            Waypoint PosA_pick: TCP in base x=15.039 y=-636.805 z=98.001 mm, rx=-1.0907 ry=1.4048 rz=-1.4136 rad; joints [-59.046, -153.942, -49.224, -157.253, 46.333, 1.224] deg
            URCap Gripper (Robotiq_Grippers, Robotiq Inc.) dataModel(position=100.0, force=30.19607843137255, speed=49.80392156862745, positionInDouble=100.0, forceInDouble=30.19607843137255, speedInDouble=49.80392156862745, slaveIds=[9], blocking=true, robotCompliant=false)
            Waypoint PosA_up: motionParameters(jointSpeed=1.047198 jointAcceleration=1.396263 cartesianSpeed=0.04 cartesianAcceleration=0.3); TCP in base x=16.801 y=-634.608 z=234.973 mm, rx=-1.0907 ry=1.4048 rz=-1.4136 rad; joints [-58.842, -146.487, -43.11, -170.828, 46.488, 1.231] deg
            Waypoint Postions_otw: motionParameters(blendRadius=0.01); TCP in base x=-10.897 y=-533.369 z=288.851 mm, rx=-1.2337 ry=1.1953 rz=-1.2073 rad; joints [-51.497, -119.089, -83.078, -158.276, 37.645, 1.224] deg
        ElseIf powder_position≟"Position2"
          MoveJ speed 60 deg/s, acceleration 80 deg/s^2 (useActiveTCP=true optimoveEnabled=false optiMoveSpeed=0.3 optiMoveAcceleration=0.09) feature=Base
            Waypoint Postions_otw: motionParameters(blendRadius=0.01); TCP in base x=-10.897 y=-533.369 z=288.851 mm, rx=-1.2337 ry=1.1953 rz=-1.2073 rad; joints [-51.497, -119.089, -83.078, -158.276, 37.645, 1.224] deg
          URCap Gripper (Robotiq_Grippers, Robotiq Inc.) dataModel(position=0.0, force=30.19607843137255, speed=49.80392156862745, positionInDouble=0.0, forceInDouble=30.19607843137255, speedInDouble=49.80392156862745, slaveIds=[9], blocking=true, robotCompliant=false)
          MoveL speed 250 mm/s, acceleration 1200 mm/s^2 (useActiveTCP=true optimoveEnabled=false optiMoveSpeed=0.3 optiMoveAcceleration=0.09) feature=Base
            Waypoint PosB_up: motionParameters(blendRadius=0.01); TCP in base x=239.473 y=-492.481 z=220.768 mm, rx=-1.2337 ry=1.1953 rz=-1.2073 rad; joints [-33.233, -137.947, -61.305, -161.095, 55.866, 1.01] deg
            Waypoint PosB_pick: TCP in base x=240.63 y=-494.559 z=96.393 mm, rx=-1.2337 ry=1.1953 rz=-1.2073 rad; joints [-33.324, -146.292, -65.182, -148.873, 55.811, 1.01] deg
            URCap Gripper (Robotiq_Grippers, Robotiq Inc.) dataModel(position=100.0, force=30.19607843137255, speed=49.80392156862745, positionInDouble=100.0, forceInDouble=30.19607843137255, speedInDouble=49.80392156862745, slaveIds=[9], blocking=true, robotCompliant=false)
            Waypoint PosB_up: motionParameters(jointSpeed=1.047198 jointAcceleration=1.396263 cartesianSpeed=0.05 cartesianAcceleration=0.4); TCP in base x=239.473 y=-492.481 z=220.768 mm, rx=-1.2337 ry=1.1953 rz=-1.2073 rad; joints [-33.233, -137.947, -61.305, -161.095, 55.866, 1.01] deg
            Waypoint Postions_otw: TCP in base x=-10.897 y=-533.369 z=288.851 mm, rx=-1.2337 ry=1.1953 rz=-1.2073 rad; joints [-51.497, -119.089, -83.078, -158.276, 37.645, 1.224] deg
        ElseIf powder_position≟"Position3"
          MoveJ speed 60 deg/s, acceleration 80 deg/s^2 (useActiveTCP=true optimoveEnabled=false optiMoveSpeed=0.3 optiMoveAcceleration=0.09) feature=Base
            Waypoint Postions_otw: motionParameters(blendRadius=0.01); TCP in base x=-10.897 y=-533.369 z=288.851 mm, rx=-1.2337 ry=1.1953 rz=-1.2073 rad; joints [-51.497, -119.089, -83.078, -158.276, 37.645, 1.224] deg
            URCap Gripper (Robotiq_Grippers, Robotiq Inc.) dataModel(position=0.0, force=30.19607843137255, speed=49.80392156862745, positionInDouble=0.0, forceInDouble=30.19607843137255, speedInDouble=49.80392156862745, slaveIds=[9], blocking=true, robotCompliant=false)
          MoveL speed 250 mm/s, acceleration 1200 mm/s^2 (useActiveTCP=true optimoveEnabled=false optiMoveSpeed=0.3 optiMoveAcceleration=0.09) feature=Base
            Waypoint PosC_up: motionParameters(blendRadius=0.01); TCP in base x=241.567 y=-359.249 z=230.261 mm, rx=-1.2337 ry=1.1953 rz=-1.2073 rad; joints [-22.674, -126.16, -80.875, -153.323, 66.473, 0.967] deg
            Waypoint PosC_pick: TCP in base x=240.634 y=-361.553 z=93.98 mm, rx=-1.2337 ry=1.1953 rz=-1.2073 rad; joints [-22.914, -136.71, -85.338, -138.313, 66.273, 0.981] deg
            URCap Gripper (Robotiq_Grippers, Robotiq Inc.) dataModel(position=100.0, force=30.19607843137255, speed=49.80392156862745, positionInDouble=100.0, forceInDouble=30.19607843137255, speedInDouble=49.80392156862745, slaveIds=[9], blocking=true, robotCompliant=false)
            Waypoint PosC_up: motionParameters(jointSpeed=1.047198 jointAcceleration=1.396263 cartesianSpeed=0.05 cartesianAcceleration=0.5); TCP in base x=241.567 y=-359.249 z=230.261 mm, rx=-1.2337 ry=1.1953 rz=-1.2073 rad; joints [-22.674, -126.16, -80.875, -153.323, 66.473, 0.967] deg
        MoveJ speed 60 deg/s, acceleration 80 deg/s^2 (useActiveTCP=true optimoveEnabled=false optiMoveSpeed=0.3 optiMoveAcceleration=0.09) feature=Base
          Waypoint Pow_decap_up: TCP in base x=-17.556 y=-367.52 z=275.835 mm, rx=-0.6056 ry=1.8925 rz=-1.8908 rad; joints [-64.584, -121.318, -81.647, -157.483, 81.325, 1.332] deg
        Set DigitalOutput pin=digital_out[5]; digitalValue=1
        Wait Sleep waitTime=0.5
        MoveL speed 50 mm/s, acceleration 500 mm/s^2 (useActiveTCP=true optimoveEnabled=false optiMoveSpeed=0.3 optiMoveAcceleration=0.09) feature=Base
          Waypoint pow_decap_place: TCP in base x=-20.433 y=-368.31 z=161.281 mm, rx=-0.6056 ry=1.8925 rz=-1.8908 rad; joints [-64.879, -129.041, -87.675, -143.733, 81.069, 1.345] deg
        Set DigitalOutput pin=digital_out[5]; digitalValue=0
        Wait Sleep waitTime=0.5
        URCap Gripper (Robotiq_Grippers, Robotiq Inc.) dataModel(position=0.0, force=30.19607843137255, speed=100.0, positionInDouble=0.0, forceInDouble=30.19607843137255, speedInDouble=100.0, slaveIds=[9], blocking=true, robotCompliant=false)
        MoveL speed 250 mm/s, acceleration 1200 mm/s^2 (useActiveTCP=true optimoveEnabled=false optiMoveSpeed=0.3 optiMoveAcceleration=0.09) feature=Base
          Waypoint Pow_decap_up: TCP in base x=-17.556 y=-367.52 z=275.835 mm, rx=-0.6056 ry=1.8925 rz=-1.8908 rad; joints [-64.584, -121.318, -81.647, -157.483, 81.325, 1.332] deg
          Waypoint Postions_otw: TCP in base x=-10.897 y=-533.369 z=288.851 mm, rx=-1.2337 ry=1.1953 rz=-1.2073 rad; joints [-51.497, -119.089, -83.078, -158.276, 37.645, 1.224] deg
        SafeHome (positionOptionType=SPEED_AND_ACCELERATION speed=1.047198 acceleration=1.396263 nextMotionTime=2)
        MoveL speed 250 mm/s, acceleration 1200 mm/s^2 (useActiveTCP=true optimoveEnabled=false optiMoveSpeed=0.3 optiMoveAcceleration=0.09) feature=Base
          Waypoint Decap_above: TCP in base x=-31.864 y=-349.975 z=288.042 mm, rx=0 ry=0 rz=0 rad; joints [-72.875, -66.865, -113.978, -89.149, 90.141, -162.862] deg
          Waypoint Decapp: TCP in base x=-31.864 y=-349.975 z=230.259 mm, rx=0 ry=0 rz=0 rad; joints [-72.901, -67.669, -121.993, -80.33, 90.142, -162.853] deg
        URCap Gripper (Robotiq_Grippers, Robotiq Inc.) dataModel(position=100.0, force=30.19607843137255, speed=50.0, positionInDouble=100.0, forceInDouble=30.19607843137255, speedInDouble=50.0, slaveIds=[9], blocking=true, robotCompliant=false)
        Folder Decap
          Action_Info := "decapping"
          Set DigitalOutput pin=GRP_3F_Enable; digitalValue=1
          Set DigitalOutput pin=GRP_3F_Decap; digitalValue=1
          Force Frame feature=Base; selection=[0, 0, 1, 0, 0, 0]; wrench=[0, 0, 2, 0, 0, 0]; limitsForce=[0.15, 0.15, 0.0005, 1.047198, 1.047198, 1.047198]; limitsMotion=[0.1, 0.1, 0.1, 0.349066, 0.349066, 0.349066]
            Script: check_decapping(offset=0.010, timeout=4.5, abort=CMD_Hold)
          Set DigitalOutput pin=GRP_3F_Decap; digitalValue=0
          Set DigitalOutput pin=GRP_3F_Enable; digitalValue=0
        MoveL speed 250 mm/s, acceleration 1200 mm/s^2 (useActiveTCP=true optimoveEnabled=false optiMoveSpeed=0.3 optiMoveAcceleration=0.09) feature=Base
          Waypoint Decap_above: TCP in base x=-31.864 y=-349.975 z=288.042 mm, rx=0 ry=0 rz=0 rad; joints [-72.875, -66.865, -113.978, -89.149, 90.141, -162.862] deg
          Waypoint Cap_above: motionParameters(blendRadius=0.05); TCP in base x=-224.192 y=-629.6 z=257.274 mm, rx=0 ry=0 rz=-1.6478 rad; joints [-98.013, -112.725, -72.795, -84.467, 90.155, -93.665] deg
          Waypoint Cap_place: TCP in base x=-224.189 y=-629.598 z=41.886 mm, rx=0 ry=0 rz=-1.6478 rad; joints [-98.043, -122.601, -91.335, -56.05, 90.142, -93.6] deg
          URCap Gripper (Robotiq_Grippers, Robotiq Inc.) dataModel(position=26.274509803921568, force=30.19607843137255, speed=30.19607843137255, positionInDouble=26.274509803921568, forceInDouble=30.19607843137255, speedInDouble=30.19607843137255, slaveIds=[9], blocking=true)
          Waypoint Cap_above: motionParameters(blendRadius=0.05); TCP in base x=-224.192 y=-629.6 z=257.274 mm, rx=0 ry=0 rz=-1.6478 rad; joints [-98.013, -112.725, -72.795, -84.467, 90.155, -93.665] deg
          SafeHome (positionOptionType=SPEED_AND_ACCELERATION speed=1.047198 acceleration=1.396263 nextMotionTime=2)
    Case (caseValue=45)
      Folder Place the decapped container- recipe
        SuppressedNode
          Script: tilt_to_home()
        SuppressedNode
          Script: tilt_send(4)
        URCap VISOR Robotic App (SensoPart VISOR Robotic, SensoPart Industriesensorik GmbH) dataModel(visorAppTemplate=1); state(isChildrenLocked=true)
          URCap Easy Pick Setup (SensoPart VISOR Robotic, SensoPart Industriesensorik GmbH) dataModel(visorId=0, visorImageAcqSetup=2, visorDetector=1, visorSetJob=true, visorOffsetSet=true, visorImageAcqSource=2, visorJobName=PoTS, visorSetupStatus=2, Pose(key=visorGripPose, Position(key=posePosition, Length(key=X value=-0.651507 unit=M), Length(key=Y value=-0.091399 unit=M), Length(key=Z value=0.249944 unit=M)), Rotation(key=poseRotation, Angle(key=RX value=-0.835678 unit=RAD), Angle(key=RY value=1.667065 unit=RAD), Angle(key=RZ value=-1.691229 unit=RAD))), Feature(key=visorImageAcqFeature name=Trigger)); state(isChildrenLocked=true)
          URCap Process (SensoPart VISOR Robotic, SensoPart Industriesensorik GmbH) dataModel(Variable(key=visorCounterVar, variable=easyPickCount_7), Variable(key=visorPartsFoundVar, variable=easyPickParts_7)); state(isChildrenLocked=true)
            URCap Image Acquisition Pose (SensoPart VISOR Robotic, SensoPart Industriesensorik GmbH) state(isChildrenLocked=true)
            URCap Object Detected (SensoPart VISOR Robotic, SensoPart Industriesensorik GmbH) state(isChildrenLocked=true)
              Folder Open Gripper
                URCap Gripper (Robotiq_Grippers, Robotiq Inc.) dataModel(position=0.0, force=30.19607843137255, speed=30.19607843137255, positionInDouble=0.0, forceInDouble=30.19607843137255, speedInDouble=30.19607843137255, slaveIds=[9], blocking=true)
                MoveL speed 250 mm/s, acceleration 1200 mm/s^2 (useActiveTCP=true optimoveEnabled=false optiMoveSpeed=0.3 optiMoveAcceleration=0.09) feature=Base
                  Waypoint OP_PowderA2: TCP in base x=9.371 y=-409.434 z=294.169 mm, rx=-0.8233 ry=1.7094 rz=-1.6983 rad; joints [-57.265, -122.586, -76.992, -161.25, 72.295, 1.124] deg; TCP offset x=0 y=0 z=161 mm, rx=3.1415 ry=0 rz=0 rad
                  Waypoint Decap_up: TCP in base x=-18.339 y=-367.674 z=249.554 mm, rx=-0.5462 ry=1.936 rz=-1.9301 rad; joints [-66.356, -123.587, -82.167, -154.733, 83.403, 1.181] deg; TCP offset x=0 y=0 z=161 mm, rx=3.1415 ry=0 rz=0 rad
                  Waypoint Decap_pick: TCP in base x=-20.429 y=-367.972 z=161.604 mm, rx=-0.5462 ry=1.936 rz=-1.9301 rad; joints [-66.558, -129.69, -86.443, -144.354, 83.231, 1.191] deg
                  URCap Gripper (Robotiq_Grippers, Robotiq Inc.) dataModel(position=100.0, force=30.19607843137255, speed=30.19607843137255, positionInDouble=100.0, forceInDouble=30.19607843137255, speedInDouble=30.19607843137255, slaveIds=[9], blocking=true, robotCompliant=false)
                  Wait Sleep waitTime=0.5
                  Set DigitalOutput pin=GRP_3F_Open; digitalValue=1
                  Waypoint Decap_up: motionParameters(jointSpeed=1.047198 jointAcceleration=1.396263 cartesianSpeed=0.1 cartesianAcceleration=0.5); TCP in base x=-18.339 y=-367.674 z=249.554 mm, rx=-0.5462 ry=1.936 rz=-1.9301 rad; joints [-66.356, -123.587, -82.167, -154.733, 83.403, 1.181] deg
                  SuppressedNode
                    Script: Motors_off()
                  Waypoint Op_PowA_wP: TCP in base x=-173.728 y=-372.934 z=295.117 mm, rx=-0.9724 ry=1.541 rz=-1.5487 rad; joints [-67.269, -106.894, -99.849, -153.52, 49.211, 1.028] deg
              URCap Approach Pose (SensoPart VISOR Robotic, SensoPart Industriesensorik GmbH) dataModel(visorOffsetZ=0.0, visorJointSpeed=25.0, visorJointAcc=30.0); state(isChildrenLocked=true)
              URCap Target Pose (SensoPart VISOR Robotic, SensoPart Industriesensorik GmbH) dataModel(visorToolSpeed=50.0, visorToolAcc=100.0); state(isChildrenLocked=true)
              Folder Close Gripper
                container_place := get_actual_tcp_pose()
                target_pose := pose_add(container_place, p[0,0,-0.12,0,0,0])
                MoveL speed 250 mm/s, acceleration 1200 mm/s^2 (useActiveTCP=true optimoveEnabled=false optiMoveSpeed=0.3 optiMoveAcceleration=0.09) feature=Base
                  Waypoint Variable (Variable): motionParameters(jointSpeed=1.047198 jointAcceleration=1.396263 cartesianSpeed=0.05 cartesianAcceleration=0.3); variable=target_pose
                URCap Gripper (Robotiq_Grippers, Robotiq Inc.) dataModel(position=0.0, force=30.19607843137255, speed=30.19607843137255, positionInDouble=0.0, forceInDouble=30.19607843137255, speedInDouble=30.19607843137255, slaveIds=[9], blocking=true)
              URCap Exit Pose (SensoPart VISOR Robotic, SensoPart Industriesensorik GmbH) dataModel(visorOffsetZ=0.0); state(isChildrenLocked=true)
            URCap No Object Detected (SensoPart VISOR Robotic, SensoPart Industriesensorik GmbH) dataModel(Variable(key=visorNoObjCountVar, variable=easyPickNoObj_7))
              Popup Message (haltProgram=false message=No weigh scale detected inputType=Text)
        place_pose := get_actual_tcp_pose()
        Script: center_pose()
        SuppressedNode
          center_tilt_pos := P_center
        MoveJ speed 60 deg/s, acceleration 80 deg/s^2 (useActiveTCP=true optimoveEnabled=false optiMoveSpeed=0.3 optiMoveAcceleration=0.09) feature=Base
          Waypoint Waypoint_1: TCP in base x=-451.049 y=-340.589 z=308.224 mm, rx=0.0971 ry=0.091 rz=-1.5784 rad; joints [-127.334, -100.578, -80.109, -94.907, 86.186, -126.663] deg
    Case (caseValue=46)
      Folder Powder dosing for recipe
        SuppressedNode
          Script: zero_scale()
        Script: send_target_info()
        Wait Sleep waitTime=0.5
        Script: send_powder_info()
        Wait Sleep waitTime=0.5
        SuppressedNode
          Folder spatula_selection test
            weight_value := get_weight()
            diff := target_weight-weight_value
            Script: scooping_init()
            Script: compute_level_percent(W_now, weight_value)
            Script: spatula = select_spatula(Pow_name, level, diff)
        URCap VISOR Robotic App (SensoPart VISOR Robotic, SensoPart Industriesensorik GmbH) dataModel(visorAppTemplate=1); state(isChildrenLocked=true)
          URCap Easy Pick Setup (SensoPart VISOR Robotic, SensoPart Industriesensorik GmbH) dataModel(visorId=0, visorSetJob=true, visorImageAcqSetup=2, visorCalibSetNo=9, visorDetector=1, visorImageAcqSource=2, visorJobName=Weight_scale, visorOffsetSet=true, visorSetupStatus=3, Pose(key=visorGripPose, Position(key=posePosition, Length(key=X value=-0.535221 unit=M), Length(key=Y value=0.017694 unit=M), Length(key=Z value=0.123958 unit=M)), Rotation(key=poseRotation, Angle(key=RX value=0.727814 unit=RAD), Angle(key=RY value=1.465761 unit=RAD), Angle(key=RZ value=-0.763944 unit=RAD))), Feature(key=visorImageAcqFeature name=Trigger)); state(isChildrenLocked=true)
          URCap Process (SensoPart VISOR Robotic, SensoPart Industriesensorik GmbH) dataModel(Variable(key=visorCounterVar, variable=easyPickCount_4), Variable(key=visorPartsFoundVar, variable=easyPickParts_4)); state(isChildrenLocked=true)
            URCap Image Acquisition Pose (SensoPart VISOR Robotic, SensoPart Industriesensorik GmbH) state(isChildrenLocked=true)
            URCap Object Detected (SensoPart VISOR Robotic, SensoPart Industriesensorik GmbH) state(isChildrenLocked=true)
              Folder Open Gripper
                Script: tare_scale()
                Wait Sleep waitTime=0.2
                weight_value := get_weight()
                Wait Sleep waitTime=0.2
                diff := target_weight-weight_value
                Script: scooping_init()
                Script: compute_level_percent(W_now, weight_value)
                Script: send_level_info()
                Script: spatula = select_spatula(Pow_name, level, diff)
                Wait Sleep waitTime=0.2
                Script: send_spatula_info()
                If spatula ≟ "spatula_L"
                  MoveJ speed 60 deg/s, acceleration 80 deg/s^2 (useActiveTCP=true optimoveEnabled=false optiMoveSpeed=0.3 optiMoveAcceleration=0.09) feature=Base
                    Waypoint Spatula_otw: TCP in base x=-38.472 y=-263.141 z=425.351 mm, rx=-0.0004 ry=-0.0001 rz=3.0344 rad; joints [-68.119, -57.773, -97.702, -114.504, 90.127, 27.957] deg
                    Waypoint pick_spat_L_abv: TCP in base x=239.059 y=-67.213 z=280.721 mm, rx=0 ry=-0.0005 rz=3.1068 rad; joints [16.774, -49.077, -122.624, -98.282, 90.162, 108.776] deg
                  MoveL speed 250 mm/s, acceleration 1200 mm/s^2 (useActiveTCP=true optimoveEnabled=false optiMoveSpeed=0.3 optiMoveAcceleration=0.09) feature=Base
                    Waypoint spat_L_pick: TCP in base x=242.469 y=-67.302 z=193.171 mm, rx=0 ry=-0.0005 rz=3.1068 rad; joints [16.429, -49.275, -135.385, -85.324, 90.17, 108.483] deg
                    URCap Gripper (Robotiq_Grippers, Robotiq Inc.) dataModel(position=100.0, force=30.0, speed=0.0, positionInDouble=100.0, forceInDouble=30.0, speedInDouble=0.0, slaveIds=[9], blocking=true)
                    Waypoint spat_L_lift: motionParameters(blendRadius=0.01); TCP in base x=245.402 y=-67.432 z=289.049 mm, rx=0 ry=-0.0005 rz=3.1068 rad; joints [16.24, -50.411, -121.005, -98.568, 90.16, 108.238] deg
                    Waypoint spat_L_side: motionParameters(blendRadius=0.01); TCP in base x=247.134 y=-17.634 z=289.063 mm, rx=0 ry=-0.0005 rz=3.1068 rad; joints [28.487, -49.174, -121.365, -99.443, 90.16, 120.484] deg
                    Waypoint spat_L_up: motionParameters(blendRadius=0.05); TCP in base x=247.136 y=-17.665 z=397.131 mm, rx=0 ry=-0.0005 rz=3.1068 rad; joints [28.565, -53.55, -103.607, -112.824, 90.132, 120.503] deg
                  MoveJ speed 60 deg/s, acceleration 80 deg/s^2 (useActiveTCP=true optimoveEnabled=false optiMoveSpeed=0.3 optiMoveAcceleration=0.09) feature=Base
                    Waypoint Spatula_otw: TCP in base x=-38.472 y=-263.141 z=425.351 mm, rx=-0.0004 ry=-0.0001 rz=3.0344 rad; joints [-68.119, -57.773, -97.702, -114.504, 90.127, 27.957] deg
                ElseIf spatula ≟"spatula_M"
                  MoveJ speed 60 deg/s, acceleration 80 deg/s^2 (useActiveTCP=true optimoveEnabled=false optiMoveSpeed=0.3 optiMoveAcceleration=0.09) feature=Base
                    Waypoint Spatula_otw: TCP in base x=-38.472 y=-263.141 z=425.351 mm, rx=-0.0004 ry=-0.0001 rz=3.0344 rad; joints [-68.119, -57.773, -97.702, -114.504, 90.127, 27.957] deg
                    Waypoint spat_M_up: motionParameters(blendRadius=0.05); TCP in base x=245.496 y=-112.113 z=420.344 mm, rx=0 ry=-0.0005 rz=3.0677 rad; joints [5.167, -58.065, -98.393, -113.528, 90.127, 99.337] deg
                  MoveL speed 250 mm/s, acceleration 1200 mm/s^2 (useActiveTCP=true optimoveEnabled=false optiMoveSpeed=0.3 optiMoveAcceleration=0.09) feature=Base
                    Waypoint spat_M_pick: TCP in base x=244.674 y=-111.985 z=192.299 mm, rx=0 ry=-0.0005 rz=3.0677 rad; joints [5.062, -53.127, -134.29, -82.569, 90.166, 99.363] deg
                    URCap Gripper (Robotiq_Grippers, Robotiq Inc.) dataModel(position=100.0, force=30.0, speed=0.0, positionInDouble=100.0, forceInDouble=30.0, speedInDouble=0.0, slaveIds=[9], blocking=true)
                    Waypoint spat_M_up: motionParameters(blendRadius=0.05); TCP in base x=245.496 y=-112.113 z=420.344 mm, rx=0 ry=-0.0005 rz=3.0677 rad; joints [5.167, -58.065, -98.393, -113.528, 90.127, 99.337] deg
                    Waypoint Spatula_otw: TCP in base x=-38.472 y=-263.141 z=425.351 mm, rx=-0.0004 ry=-0.0001 rz=3.0344 rad; joints [-68.119, -57.773, -97.702, -114.504, 90.127, 27.957] deg
                  switch_spat_M := False
                ElseIf spatula≟"spatula_S"
                  MoveJ speed 60 deg/s, acceleration 80 deg/s^2 (useActiveTCP=true optimoveEnabled=false optiMoveSpeed=0.3 optiMoveAcceleration=0.09) feature=Base
                    Waypoint Spatula_otw: TCP in base x=-38.472 y=-263.141 z=425.351 mm, rx=-0.0004 ry=-0.0001 rz=3.0344 rad; joints [-68.119, -57.773, -97.702, -114.504, 90.127, 27.957] deg
                    Waypoint spat_S_Up_9: motionParameters(blendRadius=0.05); TCP in base x=252.088 y=-159.242 z=423.282 mm, rx=0 ry=-0.0005 rz=3.0677 rad; joints [-5.618, -62.24, -96.192, -111.556, 90.127, 88.551] deg
                  MoveL speed 250 mm/s, acceleration 1200 mm/s^2 (useActiveTCP=true optimoveEnabled=false optiMoveSpeed=0.3 optiMoveAcceleration=0.09) feature=Base
                    Waypoint spat_S_Pick_5: TCP in base x=245.377 y=-158.668 z=192.286 mm, rx=0 ry=-0.0005 rz=3.0677 rad; joints [-5.78, -57.937, -132.467, -79.585, 90.161, 88.525] deg
                    URCap Gripper (Robotiq_Grippers, Robotiq Inc.) dataModel(position=100.0, force=30.0, speed=0.0, positionInDouble=100.0, forceInDouble=30.0, speedInDouble=0.0, slaveIds=[9], blocking=true)
                    Waypoint spat_S_Up_10: motionParameters(blendRadius=0.05); TCP in base x=252.088 y=-159.242 z=423.282 mm, rx=0 ry=-0.0005 rz=3.0677 rad; joints [-5.618, -62.24, -96.192, -111.556, 90.127, 88.551] deg
                    Waypoint Spatula_otw: TCP in base x=-38.472 y=-263.141 z=425.351 mm, rx=-0.0004 ry=-0.0001 rz=3.0344 rad; joints [-68.119, -57.773, -97.702, -114.504, 90.127, 27.957] deg
                  switch_spat_S := False
                ElseIf spatula≟"spatula_flat_M"
                  MoveJ speed 60 deg/s, acceleration 80 deg/s^2 (useActiveTCP=true optimoveEnabled=false optiMoveSpeed=0.3 optiMoveAcceleration=0.09) feature=Base
                    Waypoint Spatula_otw: TCP in base x=-38.472 y=-263.141 z=425.351 mm, rx=-0.0004 ry=-0.0001 rz=3.0344 rad; joints [-68.119, -57.773, -97.702, -114.504, 90.127, 27.957] deg
                    Waypoint spat_flatM_up: motionParameters(blendRadius=0.05); TCP in base x=229.023 y=-211.443 z=418.634 mm, rx=0 ry=-0.0005 rz=3.0677 rad; joints [-17.294, -63.925, -96.117, -109.949, 90.128, 76.878] deg
                  MoveL speed 250 mm/s, acceleration 1200 mm/s^2 (useActiveTCP=true optimoveEnabled=false optiMoveSpeed=0.3 optiMoveAcceleration=0.09) feature=Base
                    Waypoint spat_flatM_pick: TCP in base x=241.029 y=-208.057 z=192.271 mm, rx=0 ry=-0.0005 rz=3.0677 rad; joints [-16.075, -63.047, -130.143, -76.801, 90.154, 78.231] deg
                    URCap Gripper (Robotiq_Grippers, Robotiq Inc.) dataModel(position=100.0, force=30.0, speed=0.0, positionInDouble=100.0, forceInDouble=30.0, speedInDouble=0.0, slaveIds=[9], blocking=true, robotCompliant=false)
                    Waypoint spat_flatM_up: motionParameters(blendRadius=0.05); TCP in base x=229.023 y=-211.443 z=418.634 mm, rx=0 ry=-0.0005 rz=3.0677 rad; joints [-17.294, -63.925, -96.117, -109.949, 90.128, 76.878] deg
                    Waypoint Spatula_otw: TCP in base x=-38.472 y=-263.141 z=425.351 mm, rx=-0.0004 ry=-0.0001 rz=3.0344 rad; joints [-68.119, -57.773, -97.702, -114.504, 90.127, 27.957] deg
                  switch_spat_F_M := False
                ElseIf spatula≟"spatula_flat_S"
                  MoveJ speed 60 deg/s, acceleration 80 deg/s^2 (useActiveTCP=true optimoveEnabled=false optiMoveSpeed=0.3 optiMoveAcceleration=0.09) feature=Base
                    Waypoint Spatula_otw: TCP in base x=-38.472 y=-263.141 z=425.351 mm, rx=-0.0004 ry=-0.0001 rz=3.0344 rad; joints [-68.119, -57.773, -97.702, -114.504, 90.127, 27.957] deg
                    Waypoint spat_flatS_up: motionParameters(blendRadius=0.05); TCP in base x=237.652 y=-253.944 z=403.961 mm, rx=0 ry=-0.0005 rz=3.0677 rad; joints [-24.273, -68.411, -95.947, -105.635, 90.132, 69.906] deg
                  MoveL speed 250 mm/s, acceleration 1200 mm/s^2 (useActiveTCP=true optimoveEnabled=false optiMoveSpeed=0.3 optiMoveAcceleration=0.09) feature=Base
                    Waypoint spat_flatS_pick: TCP in base x=241.326 y=-251.726 z=192.257 mm, rx=0 ry=-0.0005 rz=3.0677 rad; joints [-23.749, -68.568, -127.154, -74.27, 90.149, 70.556] deg
                    URCap Gripper (Robotiq_Grippers, Robotiq Inc.) dataModel(position=100.0, force=30.0, speed=0.0, positionInDouble=100.0, forceInDouble=30.0, speedInDouble=0.0, slaveIds=[9], blocking=true, robotCompliant=false)
                    Waypoint spat_flatS_up: motionParameters(blendRadius=0.05); TCP in base x=237.652 y=-253.944 z=403.961 mm, rx=0 ry=-0.0005 rz=3.0677 rad; joints [-24.273, -68.411, -95.947, -105.635, 90.132, 69.906] deg
                    Waypoint Spatula_otw: TCP in base x=-38.472 y=-263.141 z=425.351 mm, rx=-0.0004 ry=-0.0001 rz=3.0344 rad; joints [-68.119, -57.773, -97.702, -114.504, 90.127, 27.957] deg
                  switch_spat_F_S := False
                weight_value := get_weight()
                Script: auto_tilt_and_scoop(W_now, target_weight, weight_value)
              URCap Approach Pose (SensoPart VISOR Robotic, SensoPart Industriesensorik GmbH) dataModel(visorJointSpeed=10.0, visorJointAcc=15.0, visorOffsetZ=-30.0); state(isChildrenLocked=true)
              URCap Target Pose (SensoPart VISOR Robotic, SensoPart Industriesensorik GmbH) dataModel(visorToolSpeed=20.0, visorToolAcc=50.0); state(isChildrenLocked=true)
              Folder Close Gripper
                dispense_pos := get_actual_tcp_pose()
                Loop While (checkContinuously=true) expression=weight_value≤target_weight
                  MoveL speed 250 mm/s, acceleration 1200 mm/s^2 (useActiveTCP=true optimoveEnabled=false optiMoveSpeed=0.3 optiMoveAcceleration=0.09) feature=Base
                    Waypoint Variable (Variable): motionParameters(jointSpeed=0.436332 jointAcceleration=0.523599 cartesianSpeed=0.1 cartesianAcceleration=0.2); variable=dispense_pos
                    Script: log_weight()
                    Wait Sleep waitTime=0.5
                    If level≥90.0
                      Script: Rotate()
                    If level≤85
                      Script: tilt_to_home()
                    Wait Sleep waitTime=0.5
                    Start_thread := True
                    vib_thread := True
                    SuppressedNode
                      tilt_angle := current_pose[5]
                    Wait Sleep waitTime=0.5
                    SuppressedNode
                      Loop While (checkContinuously=true) expression=diff>3.0
                        tilt_pose := pose_trans(get_actual_tcp_pose(), p[0, 0, 0, 0, 0, 1.0])
                        Script: movel(tilt_pose, a=0.1, v=0.1, r=0.00001)
                        tilt_pose := pose_trans(get_actual_tcp_pose(), p[0, 0, 0, 0, 0, -1.0])
                        Script: movel(tilt_pose, a=0.1, v=0.1, r=0.00001)
                    If diff ≥(target_g +(0.1*target_g))
                      tilt_pose := pose_trans(get_actual_tcp_pose(), p[0, 0, 0, 0, 0, 2.0])
                      Script: movel(tilt_pose, a=0.1, v=0.1, r=0.00001)
                    Else 
                      Loop While (checkContinuously=true) expression=weight_value≤target_weight and tilt_angle≥(-1.999) and tilt_angle≤0.5
                        current_error := target_weight-weight_value
                        Integral_error := Integral_error+current_error*dt
                        derivative := (current_error-previous_error)/dt
                        tilt_increment := (kp*current_error)+(ki*Integral_error)+(kd*derivative)
                        current_pose := get_actual_tcp_pose()
                        tilt_angle := current_pose[5]
                        tilt_pose := pose_trans(current_pose, p[0, 0, 0, 0, 0, tilt_increment])
                        Script: movel(tilt_pose, a=0.1, v=0.1, r=0.00001)
                        previous_error := current_error
                    Start_thread := False
                    SuppressedNode
                      Waypoint Waypoint_64: motionParameters(jointSpeed=1.047198 jointAcceleration=1.396263 cartesianSpeed=0.03 cartesianAcceleration=0.1 blendRadius=0.05); TCP in base x=-542.998 y=-117.021 z=221.977 mm, rx=1.8981 ry=-0.7227 rz=1.5827 rad; joints [-123.845, -120.87, -101.018, -172.406, 14.907, 127.864] deg
                    weight_value := get_weight()
                    tilt_angle := -1
                    Wait Sleep waitTime=0.5
                    vib_thread := False
                    MoveL speed 250 mm/s, acceleration 500 mm/s^2 (useActiveTCP=true optimoveEnabled=false optiMoveSpeed=0.3 optiMoveAcceleration=0.09) feature=Base
                      Waypoint Variable (Variable): variable=dispense_pos
                    Script: compute_level_percent(W_now, weight_value)
                    Script: send_level_info()
                    Script: spatula = select_spatula(Pow_name, level, diff)
                    Wait Sleep waitTime=0.2
                    SuppressedNode
                      Script: spatula = str_cat("", spatula)
                    Integral_error := 0
                    current_error := 0
                    previous_error := 0
                    Set AnalogOutput pin=analog_out[0]; analogValue=0
                    Wait Sleep waitTime=0.2
                    Script: send_spatula_info()
                    If spatula ≟ "spatula_M" and switch_spat_M≟ True
                      MoveJ speed 60 deg/s, acceleration 80 deg/s^2 (useActiveTCP=true optimoveEnabled=false optiMoveSpeed=0.3 optiMoveAcceleration=0.09) feature=Base
                        Waypoint Spatula_otw: TCP in base x=-38.472 y=-263.141 z=425.351 mm, rx=-0.0004 ry=-0.0001 rz=3.0344 rad; joints [-68.119, -57.773, -97.702, -114.504, 90.127, 27.957] deg
                        Waypoint spat_L_up: TCP in base x=247.136 y=-17.665 z=397.131 mm, rx=0 ry=-0.0005 rz=3.1068 rad; joints [28.565, -53.55, -103.607, -112.824, 90.132, 120.503] deg
                      MoveL speed 250 mm/s, acceleration 1200 mm/s^2 (useActiveTCP=true optimoveEnabled=false optiMoveSpeed=0.3 optiMoveAcceleration=0.09) feature=Base
                        Waypoint spat_L_side: TCP in base x=247.134 y=-17.634 z=289.063 mm, rx=0 ry=-0.0005 rz=3.1068 rad; joints [28.487, -49.174, -121.365, -99.443, 90.16, 120.484] deg
                        Waypoint spat_L_lift: TCP in base x=245.402 y=-67.432 z=289.049 mm, rx=0 ry=-0.0005 rz=3.1068 rad; joints [16.24, -50.411, -121.005, -98.568, 90.16, 108.238] deg
                        Waypoint spat_L_pick: TCP in base x=242.469 y=-67.302 z=193.171 mm, rx=0 ry=-0.0005 rz=3.1068 rad; joints [16.429, -49.275, -135.385, -85.324, 90.17, 108.483] deg
                        URCap Gripper (Robotiq_Grippers, Robotiq Inc.) dataModel(position=0.0, force=30.0, speed=100.0, positionInDouble=0.0, forceInDouble=30.0, speedInDouble=100.0, slaveIds=[9], blocking=true)
                        Waypoint spat_M_pick: TCP in base x=244.674 y=-111.985 z=192.299 mm, rx=0 ry=-0.0005 rz=3.0677 rad; joints [5.062, -53.127, -134.29, -82.569, 90.166, 99.363] deg
                        URCap Gripper (Robotiq_Grippers, Robotiq Inc.) dataModel(position=100.0, force=30.0, speed=0.0, positionInDouble=100.0, forceInDouble=30.0, speedInDouble=0.0, slaveIds=[9], blocking=true)
                        Waypoint spat_M_up: TCP in base x=245.496 y=-112.113 z=420.344 mm, rx=0 ry=-0.0005 rz=3.0677 rad; joints [5.167, -58.065, -98.393, -113.528, 90.127, 99.337] deg
                        Waypoint Spatula_otw: TCP in base x=-38.472 y=-263.141 z=425.351 mm, rx=-0.0004 ry=-0.0001 rz=3.0344 rad; joints [-68.119, -57.773, -97.702, -114.504, 90.127, 27.957] deg
                      switch_spat_M := False
                    ElseIf spatula ≟ "spatula_S" and switch_spat_S ≟ True
                      MoveL speed 250 mm/s, acceleration 1200 mm/s^2 (useActiveTCP=true optimoveEnabled=false optiMoveSpeed=0.3 optiMoveAcceleration=0.09) feature=Base
                        Waypoint Spatula_otw: TCP in base x=-38.472 y=-263.141 z=425.351 mm, rx=-0.0004 ry=-0.0001 rz=3.0344 rad; joints [-68.119, -57.773, -97.702, -114.504, 90.127, 27.957] deg
                        Waypoint spat_M_up: TCP in base x=245.496 y=-112.113 z=420.344 mm, rx=0 ry=-0.0005 rz=3.0677 rad; joints [5.167, -58.065, -98.393, -113.528, 90.127, 99.337] deg
                        Waypoint spat_M_pick: TCP in base x=244.674 y=-111.985 z=192.299 mm, rx=0 ry=-0.0005 rz=3.0677 rad; joints [5.062, -53.127, -134.29, -82.569, 90.166, 99.363] deg
                        URCap Gripper (Robotiq_Grippers, Robotiq Inc.) dataModel(position=0.0, force=30.19607843137255, speed=100.0, positionInDouble=0.0, forceInDouble=30.19607843137255, speedInDouble=100.0, slaveIds=[9], blocking=true)
                        Waypoint spat_S_pick: TCP in base x=238.159 y=-157.927 z=192.632 mm, rx=0 ry=-0.0005 rz=3.0677 rad; joints [-5.778, -56.616, -132.95, -80.422, 90.162, 88.526] deg
                        URCap Gripper (Robotiq_Grippers, Robotiq Inc.) dataModel(position=100.0, force=30.19607843137255, speed=0.0, positionInDouble=100.0, forceInDouble=30.19607843137255, speedInDouble=0.0, slaveIds=[9], blocking=true)
                        Waypoint spat_S_up: TCP in base x=244.261 y=-164.467 z=417.088 mm, rx=0 ry=-0.0005 rz=3.0677 rad; joints [-6.934, -61.411, -97.537, -111.041, 90.129, 87.239] deg
                        Waypoint Spatula_otw: TCP in base x=-38.472 y=-263.141 z=425.351 mm, rx=-0.0004 ry=-0.0001 rz=3.0344 rad; joints [-68.119, -57.773, -97.702, -114.504, 90.127, 27.957] deg
                      switch_spat_S := False
                    ElseIf spatula≟"spatula_flat_S"  and switch_spat_F_S ≟ True
                      MoveL speed 250 mm/s, acceleration 1200 mm/s^2 (useActiveTCP=true optimoveEnabled=false optiMoveSpeed=0.3 optiMoveAcceleration=0.09) feature=Base
                        Waypoint Spatula_otw: TCP in base x=-38.472 y=-263.141 z=425.351 mm, rx=-0.0004 ry=-0.0001 rz=3.0344 rad; joints [-68.119, -57.773, -97.702, -114.504, 90.127, 27.957] deg
                        Waypoint spat_flatM_up: TCP in base x=229.023 y=-211.443 z=418.634 mm, rx=0 ry=-0.0005 rz=3.0677 rad; joints [-17.294, -63.925, -96.117, -109.949, 90.128, 76.878] deg
                        Waypoint spat_flatM_pick: TCP in base x=241.029 y=-208.057 z=192.271 mm, rx=0 ry=-0.0005 rz=3.0677 rad; joints [-16.075, -63.047, -130.143, -76.801, 90.154, 78.231] deg
                        URCap Gripper (Robotiq_Grippers, Robotiq Inc.) dataModel(position=0.0, force=30.0, speed=0.0, positionInDouble=0.0, forceInDouble=30.0, speedInDouble=0.0, slaveIds=[9], blocking=true, robotCompliant=false)
                        Waypoint spat_flatS_pick: TCP in base x=241.326 y=-251.726 z=192.257 mm, rx=0 ry=-0.0005 rz=3.0677 rad; joints [-23.749, -68.568, -127.154, -74.27, 90.149, 70.556] deg
                        URCap Gripper (Robotiq_Grippers, Robotiq Inc.) dataModel(position=100.0, force=30.0, speed=0.0, positionInDouble=100.0, forceInDouble=30.0, speedInDouble=0.0, slaveIds=[9], blocking=true, robotCompliant=false)
                        Waypoint spat_flatS_up: TCP in base x=237.652 y=-253.944 z=403.961 mm, rx=0 ry=-0.0005 rz=3.0677 rad; joints [-24.273, -68.411, -95.947, -105.635, 90.132, 69.906] deg
                        Waypoint Spatula_otw: TCP in base x=-38.472 y=-263.141 z=425.351 mm, rx=-0.0004 ry=-0.0001 rz=3.0344 rad; joints [-68.119, -57.773, -97.702, -114.504, 90.127, 27.957] deg
                      switch_spat_F_S := False
                    Script: auto_tilt_and_scoop(W_now, target_weight, weight_value)
                    Wait Sleep waitTime=0.5
                Start_thread := False
                Wait Sleep waitTime=0.5
                vib_thread := False
                SuppressedNode
                  Script: Rotate()
              URCap Exit Pose (SensoPart VISOR Robotic, SensoPart Industriesensorik GmbH) dataModel(visorOffsetZ=0.0); state(isChildrenLocked=true)
            URCap No Object Detected (SensoPart VISOR Robotic, SensoPart Industriesensorik GmbH) dataModel(Variable(key=visorNoObjCountVar, variable=easyPickNoObj_4))
              Popup Message (haltProgram=false message=No weigh scale detected inputType=Text)
        SuppressedNode
          Task := "Dosing"
        SuppressedNode
          Script: scooping_init()
        MoveJ speed 60 deg/s, acceleration 80 deg/s^2 (useActiveTCP=true optimoveEnabled=false optiMoveSpeed=0.3 optiMoveAcceleration=0.09) feature=Base
          Waypoint Variable (Variable): motionParameters(jointSpeed=0.436332 jointAcceleration=0.523599 cartesianSpeed=0.1 cartesianAcceleration=0.2); variable=dispense_pos
        weight_value := get_weight()
        Script: after_scoop()
        If spatula≟"spatula_M"
          MoveJ speed 60 deg/s, acceleration 80 deg/s^2 (useActiveTCP=true optimoveEnabled=false optiMoveSpeed=0.3 optiMoveAcceleration=0.09) feature=Base
            Waypoint Spatula_otw: TCP in base x=-38.472 y=-263.141 z=425.351 mm, rx=-0.0004 ry=-0.0001 rz=3.0344 rad; joints [-68.119, -57.773, -97.702, -114.504, 90.127, 27.957] deg
            Waypoint spat_M_up: TCP in base x=245.496 y=-112.113 z=420.344 mm, rx=0 ry=-0.0005 rz=3.0677 rad; joints [5.167, -58.065, -98.393, -113.528, 90.127, 99.337] deg
          MoveL speed 250 mm/s, acceleration 1200 mm/s^2 (useActiveTCP=true optimoveEnabled=false optiMoveSpeed=0.3 optiMoveAcceleration=0.09) feature=Base
            Waypoint spat_M_pick: TCP in base x=244.674 y=-111.985 z=192.299 mm, rx=0 ry=-0.0005 rz=3.0677 rad; joints [5.062, -53.127, -134.29, -82.569, 90.166, 99.363] deg
            URCap Gripper (Robotiq_Grippers, Robotiq Inc.) dataModel(position=0.0, force=30.19607843137255, speed=50.0, positionInDouble=0.0, forceInDouble=30.19607843137255, speedInDouble=50.0, slaveIds=[9], blocking=true, robotCompliant=false)
            Waypoint spat_M_up: TCP in base x=245.496 y=-112.113 z=420.344 mm, rx=0 ry=-0.0005 rz=3.0677 rad; joints [5.167, -58.065, -98.393, -113.528, 90.127, 99.337] deg
          SafeHome (positionOptionType=SPEED_AND_ACCELERATION speed=1.047198 acceleration=1.396263 nextMotionTime=2)
        ElseIf spatula≟"spatula_flat_S"
          MoveJ speed 60 deg/s, acceleration 80 deg/s^2 (useActiveTCP=true optimoveEnabled=false optiMoveSpeed=0.3 optiMoveAcceleration=0.09) feature=Base
            Waypoint Spatula_otw: TCP in base x=-38.472 y=-263.141 z=425.351 mm, rx=-0.0004 ry=-0.0001 rz=3.0344 rad; joints [-68.119, -57.773, -97.702, -114.504, 90.127, 27.957] deg
            Waypoint spat_flatS_up: TCP in base x=237.652 y=-253.944 z=403.961 mm, rx=0 ry=-0.0005 rz=3.0677 rad; joints [-24.273, -68.411, -95.947, -105.635, 90.132, 69.906] deg
          MoveL speed 250 mm/s, acceleration 1200 mm/s^2 (useActiveTCP=true optimoveEnabled=false optiMoveSpeed=0.3 optiMoveAcceleration=0.09) feature=Base
            Waypoint spat_flatS_pick: TCP in base x=241.326 y=-251.726 z=192.257 mm, rx=0 ry=-0.0005 rz=3.0677 rad; joints [-23.749, -68.568, -127.154, -74.27, 90.149, 70.556] deg
            URCap Gripper (Robotiq_Grippers, Robotiq Inc.) dataModel(position=0.0, force=30.19607843137255, speed=50.0, positionInDouble=0.0, forceInDouble=30.19607843137255, speedInDouble=50.0, slaveIds=[9], blocking=true, robotCompliant=false)
            Waypoint spat_flatS_up: TCP in base x=237.652 y=-253.944 z=403.961 mm, rx=0 ry=-0.0005 rz=3.0677 rad; joints [-24.273, -68.411, -95.947, -105.635, 90.132, 69.906] deg
          SafeHome (positionOptionType=SPEED_AND_ACCELERATION speed=1.047198 acceleration=1.396263 nextMotionTime=2)
        Folder Pick container from PoTS
          cont_place_offs := pose_add(container_place, p[0.05,0,0,0,0,0])
          MoveJ speed 60 deg/s, acceleration 80 deg/s^2 (useActiveTCP=true optimoveEnabled=false optiMoveSpeed=0.3 optiMoveAcceleration=0.09) feature=Base
            Waypoint Variable (Variable): variable=cont_place_offs
            Waypoint Variable (Variable): variable=container_place
          MoveL speed 250 mm/s, acceleration 1200 mm/s^2 (useActiveTCP=true optimoveEnabled=false optiMoveSpeed=0.3 optiMoveAcceleration=0.09) feature=Base
            Waypoint Variable (Variable): variable=target_pose
            URCap Gripper (Robotiq_Grippers, Robotiq Inc.) dataModel(position=100.0, force=30.0, speed=30.0, positionInDouble=100.0, forceInDouble=30.0, speedInDouble=30.0, slaveIds=[9], blocking=true, robotCompliant=false)
            Waypoint Variable (Variable): motionParameters(jointSpeed=1.047198 jointAcceleration=1.396263 cartesianSpeed=0.1 cartesianAcceleration=0.6); variable=container_place
        SuppressedNode
          powder_position := "Position2"
        Folder Place Powder container back to holder
          If powder_position ≟ "Position1"
            MoveL speed 250 mm/s, acceleration 1200 mm/s^2 (useActiveTCP=true optimoveEnabled=false optiMoveSpeed=0.3 optiMoveAcceleration=0.09) feature=Base
              Waypoint Postions_otw: motionParameters(blendRadius=0.01); TCP in base x=-10.897 y=-533.369 z=288.851 mm, rx=-1.2337 ry=1.1953 rz=-1.2073 rad; joints [-51.497, -119.089, -83.078, -158.276, 37.645, 1.224] deg
            MoveL speed 250 mm/s, acceleration 1200 mm/s^2 (useActiveTCP=true optimoveEnabled=false optiMoveSpeed=0.3 optiMoveAcceleration=0.09) feature=Base
              Waypoint PosA_up: TCP in base x=16.801 y=-634.608 z=234.973 mm, rx=-1.0907 ry=1.4048 rz=-1.4136 rad; joints [-58.842, -146.487, -43.11, -170.828, 46.488, 1.231] deg
              Waypoint PosA_pick: motionParameters(jointSpeed=1.047198 jointAcceleration=1.396263 cartesianSpeed=0.05 cartesianAcceleration=0.3); TCP in base x=15.039 y=-636.805 z=98.001 mm, rx=-1.0907 ry=1.4048 rz=-1.4136 rad; joints [-59.046, -153.942, -49.224, -157.253, 46.333, 1.224] deg
              URCap Gripper (Robotiq_Grippers, Robotiq Inc.) dataModel(position=0.0, force=30.19607843137255, speed=50.0, positionInDouble=0.0, forceInDouble=30.19607843137255, speedInDouble=50.0, slaveIds=[9], blocking=true, robotCompliant=false)
              Waypoint PosA_up: TCP in base x=16.801 y=-634.608 z=234.973 mm, rx=-1.0907 ry=1.4048 rz=-1.4136 rad; joints [-58.842, -146.487, -43.11, -170.828, 46.488, 1.231] deg
              Waypoint Postions_otw: motionParameters(blendRadius=0.05); TCP in base x=-10.897 y=-533.369 z=288.851 mm, rx=-1.2337 ry=1.1953 rz=-1.2073 rad; joints [-51.497, -119.089, -83.078, -158.276, 37.645, 1.224] deg
          ElseIf powder_position≟"Position2"
            MoveL speed 250 mm/s, acceleration 1200 mm/s^2 (useActiveTCP=true optimoveEnabled=false optiMoveSpeed=0.3 optiMoveAcceleration=0.09) feature=Base
              Waypoint Postions_otw: motionParameters(blendRadius=0.01); TCP in base x=-10.897 y=-533.369 z=288.851 mm, rx=-1.2337 ry=1.1953 rz=-1.2073 rad; joints [-51.497, -119.089, -83.078, -158.276, 37.645, 1.224] deg
            MoveL speed 250 mm/s, acceleration 1200 mm/s^2 (useActiveTCP=true optimoveEnabled=false optiMoveSpeed=0.3 optiMoveAcceleration=0.09) feature=Base
              Waypoint PosB_up: motionParameters(blendRadius=0.01); TCP in base x=239.473 y=-492.481 z=220.768 mm, rx=-1.2337 ry=1.1953 rz=-1.2073 rad; joints [-33.233, -137.947, -61.305, -161.095, 55.866, 1.01] deg
              Waypoint PosB_pick: motionParameters(jointSpeed=1.047198 jointAcceleration=1.396263 cartesianSpeed=0.05 cartesianAcceleration=0.3); TCP in base x=240.63 y=-494.559 z=96.393 mm, rx=-1.2337 ry=1.1953 rz=-1.2073 rad; joints [-33.324, -146.292, -65.182, -148.873, 55.811, 1.01] deg
              URCap Gripper (Robotiq_Grippers, Robotiq Inc.) dataModel(position=0.0, force=30.19607843137255, speed=50.0, positionInDouble=0.0, forceInDouble=30.19607843137255, speedInDouble=50.0, slaveIds=[9], blocking=true, robotCompliant=false)
              Waypoint PosB_up: TCP in base x=239.473 y=-492.481 z=220.768 mm, rx=-1.2337 ry=1.1953 rz=-1.2073 rad; joints [-33.233, -137.947, -61.305, -161.095, 55.866, 1.01] deg
              Waypoint Postions_otw: motionParameters(blendRadius=0.05); TCP in base x=-10.897 y=-533.369 z=288.851 mm, rx=-1.2337 ry=1.1953 rz=-1.2073 rad; joints [-51.497, -119.089, -83.078, -158.276, 37.645, 1.224] deg
          ElseIf powder_position≟"Position3"
            MoveL speed 250 mm/s, acceleration 1200 mm/s^2 (useActiveTCP=true optimoveEnabled=false optiMoveSpeed=0.3 optiMoveAcceleration=0.09) feature=Base
              Waypoint Postions_otw: motionParameters(blendRadius=0.01); TCP in base x=-10.897 y=-533.369 z=288.851 mm, rx=-1.2337 ry=1.1953 rz=-1.2073 rad; joints [-51.497, -119.089, -83.078, -158.276, 37.645, 1.224] deg
            MoveL speed 250 mm/s, acceleration 1200 mm/s^2 (useActiveTCP=true optimoveEnabled=false optiMoveSpeed=0.3 optiMoveAcceleration=0.09) feature=Base
              Waypoint PosC_up: motionParameters(blendRadius=0.01); TCP in base x=241.567 y=-359.249 z=230.261 mm, rx=-1.2337 ry=1.1953 rz=-1.2073 rad; joints [-22.674, -126.16, -80.875, -153.323, 66.473, 0.967] deg
              Waypoint PosC_pick: motionParameters(jointSpeed=1.047198 jointAcceleration=1.396263 cartesianSpeed=0.05 cartesianAcceleration=0.3); TCP in base x=240.634 y=-361.553 z=93.98 mm, rx=-1.2337 ry=1.1953 rz=-1.2073 rad; joints [-22.914, -136.71, -85.338, -138.313, 66.273, 0.981] deg
              URCap Gripper (Robotiq_Grippers, Robotiq Inc.) dataModel(position=0.0, force=30.19607843137255, speed=50.0, positionInDouble=0.0, forceInDouble=30.19607843137255, speedInDouble=50.0, slaveIds=[9], blocking=true, robotCompliant=false)
              Waypoint PosC_up: TCP in base x=241.567 y=-359.249 z=230.261 mm, rx=-1.2337 ry=1.1953 rz=-1.2073 rad; joints [-22.674, -126.16, -80.875, -153.323, 66.473, 0.967] deg
              Waypoint Postions_otw: motionParameters(blendRadius=0.05); TCP in base x=-10.897 y=-533.369 z=288.851 mm, rx=-1.2337 ry=1.1953 rz=-1.2073 rad; joints [-51.497, -119.089, -83.078, -158.276, 37.645, 1.224] deg
        MoveJ speed 60 deg/s, acceleration 80 deg/s^2 (useActiveTCP=true optimoveEnabled=false optiMoveSpeed=0.3 optiMoveAcceleration=0.09) feature=Base
          Waypoint Cap_above: motionParameters(blendRadius=0.05); TCP in base x=-224.192 y=-629.6 z=257.274 mm, rx=0 ry=0 rz=-1.6478 rad; joints [-98.013, -112.725, -72.795, -84.467, 90.155, -93.665] deg
        MoveL speed 250 mm/s, acceleration 1200 mm/s^2 (useActiveTCP=true optimoveEnabled=false optiMoveSpeed=0.3 optiMoveAcceleration=0.09) feature=Base
          Waypoint Cap_place: TCP in base x=-224.189 y=-629.598 z=41.886 mm, rx=0 ry=0 rz=-1.6478 rad; joints [-98.043, -122.601, -91.335, -56.05, 90.142, -93.6] deg
          URCap Gripper (Robotiq_Grippers, Robotiq Inc.) dataModel(position=100.0, force=30.0, speed=30.0, positionInDouble=100.0, forceInDouble=30.0, speedInDouble=30.0, slaveIds=[9], blocking=true, robotCompliant=false)
          Waypoint Cap_above: motionParameters(blendRadius=0.05); TCP in base x=-224.192 y=-629.6 z=257.274 mm, rx=0 ry=0 rz=-1.6478 rad; joints [-98.013, -112.725, -72.795, -84.467, 90.155, -93.665] deg
        Folder Cap the container
          If powder_position ≟ "Position1"
            MoveJ speed 60 deg/s, acceleration 80 deg/s^2 (useActiveTCP=true optimoveEnabled=false optiMoveSpeed=0.3 optiMoveAcceleration=0.09) feature=Base
              Waypoint Cap_Pos1_up: TCP in base x=-9.205 y=-630.415 z=209.553 mm, rx=0 ry=0 rz=-1.6478 rad; joints [-78.565, -108.612, -85.584, -75.789, 90.15, -74.174] deg
            MoveL speed 250 mm/s, acceleration 1200 mm/s^2 (useActiveTCP=true optimoveEnabled=false optiMoveSpeed=0.3 optiMoveAcceleration=0.09) feature=Base
              Waypoint Cap_pos1: motionParameters(jointSpeed=1.047198 jointAcceleration=1.396263 cartesianSpeed=0.05 cartesianAcceleration=0.3); TCP in base x=-9.203 y=-630.421 z=169.124 mm, rx=0 ry=0 rz=-1.6478 rad; joints [-78.572, -110.201, -89.57, -70.215, 90.147, -74.162] deg
          ElseIf powder_position≟"Position2"
            MoveJ speed 60 deg/s, acceleration 80 deg/s^2 (useActiveTCP=true optimoveEnabled=false optiMoveSpeed=0.3 optiMoveAcceleration=0.09) feature=Base
              Waypoint Cap_Pos2_up: TCP in base x=211.716 y=-494.058 z=215.28 mm, rx=0 ry=0 rz=-1.6478 rad; joints [-52.398, -95.953, -100.395, -73.635, 90.139, -47.972] deg
            MoveL speed 50 mm/s, acceleration 300 mm/s^2 (useActiveTCP=true optimoveEnabled=false optiMoveSpeed=0.3 optiMoveAcceleration=0.09) feature=Base
              Waypoint Cap_Pos2: TCP in base x=212.49 y=-496.567 z=174.148 mm, rx=0 ry=0 rz=-1.6478 rad; joints [-52.507, -98.18, -104.219, -67.583, 90.135, -48.061] deg
          ElseIf powder_position≟"Position3"
            MoveJ speed 60 deg/s, acceleration 80 deg/s^2 (useActiveTCP=true optimoveEnabled=false optiMoveSpeed=0.3 optiMoveAcceleration=0.09) feature=Base
              Waypoint Cap_Pos3_up: TCP in base x=215.414 y=-362.498 z=204.705 mm, rx=0 ry=0 rz=-1.6478 rad; joints [-40.834, -79.894, -117.409, -72.679, 90.135, -36.369] deg
            MoveL speed 50 mm/s, acceleration 300 mm/s^2 (useActiveTCP=true optimoveEnabled=false optiMoveSpeed=0.3 optiMoveAcceleration=0.09) feature=Base
              Waypoint Cap_pos3: TCP in base x=215.415 y=-362.498 z=173.969 mm, rx=0 ry=0 rz=-1.6478 rad; joints [-40.844, -81.499, -120.873, -67.609, 90.131, -36.361] deg
          Folder Capping motion
            URCap Gripper (Robotiq_Grippers, Robotiq Inc.) dataModel(position=43.04106548279689, force=30.19607843137255, speed=30.19607843137255, positionInDouble=43.04106548279689, forceInDouble=30.19607843137255, speedInDouble=30.19607843137255, slaveIds=[9], blocking=true, robotCompliant=false)
            Loop Counting (count=2) loopVariable(name=Loop_7)
              SuppressedNode
                MoveL speed 250 mm/s, acceleration 1200 mm/s^2 (useActiveTCP=true optimoveEnabled=false optiMoveSpeed=0.3 optiMoveAcceleration=0.09) feature=Base
                  Waypoint Waypoint_4: TCP in base x=-9.21 y=-630.419 z=169.124 mm, rx=0 ry=0.0001 rz=2.738 rad; joints [-78.569, -110.197, -89.576, -70.207, 90.138, 34.552] deg
                  URCap Gripper (Robotiq_Grippers, Robotiq Inc.) dataModel(position=33.9400665926748, force=30.0, speed=30.0, positionInDouble=33.9400665926748, forceInDouble=30.0, speedInDouble=30.0, slaveIds=[9], blocking=true, robotCompliant=false)
                  Waypoint Waypoint_6: TCP in base x=-9.203 y=-630.421 z=169.124 mm, rx=-0.0001 ry=0 rz=-0.5349 rad; joints [-78.571, -110.201, -89.568, -70.218, 90.143, -137.928] deg
                  SuppressedNode
                    URCap Gripper (Robotiq_Grippers, Robotiq Inc.) dataModel(position=52.14206437291897, force=30.0, speed=30.0, positionInDouble=52.14206437291897, forceInDouble=30.0, speedInDouble=30.0, slaveIds=[9], blocking=true, robotCompliant=false)
              Cap_CW := pose_add(get_actual_tcp_pose(), p[0,0,0,0,0,2.2])
              MoveL speed 250 mm/s, acceleration 1200 mm/s^2 (useActiveTCP=true optimoveEnabled=false optiMoveSpeed=0.3 optiMoveAcceleration=0.09) feature=Base
                Waypoint Variable (Variable): variable(name=Cap_CW)
              URCap Gripper (Robotiq_Grippers, Robotiq Inc.) dataModel(position=52.14206437291897, force=30.0, speed=30.0, positionInDouble=52.14206437291897, forceInDouble=30.0, speedInDouble=30.0, slaveIds=[9], blocking=true, robotCompliant=false)
              Cap_CCW := pose_add(get_actual_tcp_pose(), p[0,0,0,0,0,-2.2])
              MoveL speed 250 mm/s, acceleration 1200 mm/s^2 (useActiveTCP=true optimoveEnabled=false optiMoveSpeed=0.3 optiMoveAcceleration=0.09) feature=Base
                Waypoint Variable (Variable): variable(name=Cap_CCW)
              URCap Gripper (Robotiq_Grippers, Robotiq Inc.) dataModel(position=43.04106548279689, force=30.19607843137255, speed=30.19607843137255, positionInDouble=43.04106548279689, forceInDouble=30.19607843137255, speedInDouble=30.19607843137255, slaveIds=[9], blocking=true, robotCompliant=false)
            URCap Gripper (Robotiq_Grippers, Robotiq Inc.) dataModel(position=0.0, force=30.0, speed=30.0, positionInDouble=0.0, forceInDouble=30.0, speedInDouble=30.0, slaveIds=[9], blocking=true, robotCompliant=false)
            after_capping := pose_add(get_actual_tcp_pose(), p[0,0,0.05,0,0,0])
            MoveL speed 250 mm/s, acceleration 1200 mm/s^2 (useActiveTCP=true optimoveEnabled=false optiMoveSpeed=0.3 optiMoveAcceleration=0.09) feature=Base
              Waypoint Variable (Variable): variable(name=after_capping)
            SafeHome (positionOptionType=SPEED_AND_ACCELERATION speed=1.047198 acceleration=1.396263 nextMotionTime=2)
    Case (caseValue=47)
      Folder Pick containers
        URCap VISOR Robotic App (SensoPart VISOR Robotic, SensoPart Industriesensorik GmbH) dataModel(visorAppTemplate=1); state(isChildrenLocked=true)
          URCap Easy Pick Setup (SensoPart VISOR Robotic, SensoPart Industriesensorik GmbH) dataModel(visorId=0, visorSetJob=true, visorJobName=Containers_pick, visorImageAcqSetup=2, visorImageAcqSource=2, visorDetector=1, visorOffsetSet=true, visorSetupStatus=3, Pose(key=visorGripPose, Position(key=posePosition, Length(key=X value=-0.550589 unit=M), Length(key=Y value=0.42966 unit=M), Length(key=Z value=-0.073092 unit=M)), Rotation(key=poseRotation, Angle(key=RX value=-0.287411 unit=RAD), Angle(key=RY value=2.087623 unit=RAD), Angle(key=RZ value=-2.089777 unit=RAD))), Feature(key=visorImageAcqFeature name=Trigger)); state(isChildrenLocked=true)
          URCap Process (SensoPart VISOR Robotic, SensoPart Industriesensorik GmbH) dataModel(Variable(key=visorCounterVar, variable(name=easyPickCount_9, initializeExpression=0)), Variable(key=visorPartsFoundVar, variable(name=easyPickParts_9, initializeExpression=0))); state(isChildrenLocked=true)
            URCap Image Acquisition Pose (SensoPart VISOR Robotic, SensoPart Industriesensorik GmbH) state(isChildrenLocked=true)
            URCap Object Detected (SensoPart VISOR Robotic, SensoPart Industriesensorik GmbH) state(isChildrenLocked=true)
              Folder Open Gripper
                URCap Gripper (Robotiq_Grippers, Robotiq Inc.) dataModel(position=0.0, force=30.19607843137255, speed=30.19607843137255, positionInDouble=0.0, forceInDouble=30.19607843137255, speedInDouble=30.19607843137255, slaveIds=[9], blocking=true, robotCompliant=false)
                MoveJ speed 60 deg/s, acceleration 80 deg/s^2 (useActiveTCP=true optimoveEnabled=false optiMoveSpeed=0.3 optiMoveAcceleration=0.09) feature=Base
                  Waypoint pick_cont_otw: TCP in base x=-479.451 y=284.141 z=125.27 mm, rx=-0.2768 ry=2.0984 rz=-2.1213 rad; joints [-165.671, -112.009, -127.874, -95.426, 1.192, -23.029] deg
              URCap Approach Pose (SensoPart VISOR Robotic, SensoPart Industriesensorik GmbH) dataModel(visorOffsetZ=-50.0); state(isChildrenLocked=true)
              URCap Target Pose (SensoPart VISOR Robotic, SensoPart Industriesensorik GmbH) dataModel(visorMotionType=1); state(isChildrenLocked=true)
              Folder Close Gripper
                URCap Gripper (Robotiq_Grippers, Robotiq Inc.) dataModel(position=100.0, force=30.19607843137255, speed=30.19607843137255, positionInDouble=100.0, forceInDouble=30.19607843137255, speedInDouble=30.19607843137255, slaveIds=[9], blocking=true, robotCompliant=false)
              URCap Exit Pose (SensoPart VISOR Robotic, SensoPart Industriesensorik GmbH) dataModel(visorOffsetZ=0.0, visorMotionType=1); state(isChildrenLocked=true)
            URCap No Object Detected (SensoPart VISOR Robotic, SensoPart Industriesensorik GmbH) dataModel(Variable(key=visorNoObjCountVar, variable(name=easyPickNoObj_9, initializeExpression=0)))
              Popup Message (haltProgram=false message=No container detected inputType=Text)
        MoveJ speed 60 deg/s, acceleration 80 deg/s^2 (useActiveTCP=true optimoveEnabled=false optiMoveSpeed=0.3 optiMoveAcceleration=0.09) feature=Base
          Waypoint Powder_wayp1: TCP in base x=-472.821 y=292.44 z=207.418 mm, rx=-0.1378 ry=2.1773 rz=-2.152 rad; joints [-166.796, -109, -112.802, -143.26, 6.548, 5.495] deg
        If powder_position ≟ "Position1"
          MoveJ speed 60 deg/s, acceleration 80 deg/s^2 (useActiveTCP=true optimoveEnabled=false optiMoveSpeed=0.3 optiMoveAcceleration=0.09) feature=Base
            Waypoint Postions_otw: motionParameters(blendRadius=0.01); TCP in base x=-10.897 y=-533.369 z=288.851 mm, rx=-1.2337 ry=1.1953 rz=-1.2073 rad; joints [-51.497, -119.089, -83.078, -158.276, 37.645, 1.224] deg
          MoveL speed 250 mm/s, acceleration 1200 mm/s^2 (useActiveTCP=true optimoveEnabled=false optiMoveSpeed=0.3 optiMoveAcceleration=0.09) feature=Base
            Waypoint PosA_up: TCP in base x=16.801 y=-634.608 z=234.973 mm, rx=-1.0907 ry=1.4048 rz=-1.4136 rad; joints [-58.842, -146.487, -43.11, -170.828, 46.488, 1.231] deg
            Waypoint PosA_pick: motionParameters(jointSpeed=1.047198 jointAcceleration=1.396263 cartesianSpeed=0.05 cartesianAcceleration=0.3); TCP in base x=15.039 y=-636.805 z=98.001 mm, rx=-1.0907 ry=1.4048 rz=-1.4136 rad; joints [-59.046, -153.942, -49.224, -157.253, 46.333, 1.224] deg
            URCap Gripper (Robotiq_Grippers, Robotiq Inc.) dataModel(position=0.0, force=30.19607843137255, speed=30.19607843137255, positionInDouble=0.0, forceInDouble=30.19607843137255, speedInDouble=30.19607843137255, slaveIds=[9], blocking=true, robotCompliant=false)
            Waypoint PosA_up: TCP in base x=16.801 y=-634.608 z=234.973 mm, rx=-1.0907 ry=1.4048 rz=-1.4136 rad; joints [-58.842, -146.487, -43.11, -170.828, 46.488, 1.231] deg
            Waypoint Postions_otw: motionParameters(blendRadius=0.01); TCP in base x=-10.897 y=-533.369 z=288.851 mm, rx=-1.2337 ry=1.1953 rz=-1.2073 rad; joints [-51.497, -119.089, -83.078, -158.276, 37.645, 1.224] deg
          powder_position := "Position2"
          SafeHome (positionOptionType=SPEED_AND_ACCELERATION speed=1.047198 acceleration=1.396263 nextMotionTime=2)
          Num_cont_picked := Num_cont_picked+1
        ElseIf powder_position≟"Position2"
          MoveJ speed 60 deg/s, acceleration 80 deg/s^2 (useActiveTCP=true optimoveEnabled=false optiMoveSpeed=0.3 optiMoveAcceleration=0.09) feature=Base
            Waypoint Postions_otw: motionParameters(blendRadius=0.01); TCP in base x=-10.897 y=-533.369 z=288.851 mm, rx=-1.2337 ry=1.1953 rz=-1.2073 rad; joints [-51.497, -119.089, -83.078, -158.276, 37.645, 1.224] deg
          MoveL speed 250 mm/s, acceleration 1200 mm/s^2 (useActiveTCP=true optimoveEnabled=false optiMoveSpeed=0.3 optiMoveAcceleration=0.09) feature=Base
            Waypoint PosB_up: motionParameters(blendRadius=0.01); TCP in base x=239.473 y=-492.481 z=220.768 mm, rx=-1.2337 ry=1.1953 rz=-1.2073 rad; joints [-33.233, -137.947, -61.305, -161.095, 55.866, 1.01] deg
            Waypoint PosB_pick: motionParameters(jointSpeed=1.047198 jointAcceleration=1.396263 cartesianSpeed=0.05 cartesianAcceleration=0.3); TCP in base x=240.63 y=-494.559 z=96.393 mm, rx=-1.2337 ry=1.1953 rz=-1.2073 rad; joints [-33.324, -146.292, -65.182, -148.873, 55.811, 1.01] deg
            URCap Gripper (Robotiq_Grippers, Robotiq Inc.) dataModel(position=0.0, force=30.19607843137255, speed=30.19607843137255, positionInDouble=0.0, forceInDouble=30.19607843137255, speedInDouble=30.19607843137255, slaveIds=[9], blocking=true, robotCompliant=false)
            Waypoint PosB_up: TCP in base x=239.473 y=-492.481 z=220.768 mm, rx=-1.2337 ry=1.1953 rz=-1.2073 rad; joints [-33.233, -137.947, -61.305, -161.095, 55.866, 1.01] deg
            Waypoint Postions_otw: TCP in base x=-10.897 y=-533.369 z=288.851 mm, rx=-1.2337 ry=1.1953 rz=-1.2073 rad; joints [-51.497, -119.089, -83.078, -158.276, 37.645, 1.224] deg
          powder_position := "Position3"
          SafeHome (positionOptionType=SPEED_AND_ACCELERATION speed=1.047198 acceleration=1.396263 nextMotionTime=2)
          Num_cont_picked := Num_cont_picked+1
        ElseIf powder_position≟"Position3"
          MoveJ speed 60 deg/s, acceleration 80 deg/s^2 (useActiveTCP=true optimoveEnabled=false optiMoveSpeed=0.3 optiMoveAcceleration=0.09) feature=Base
            Waypoint Postions_otw: motionParameters(blendRadius=0.01); TCP in base x=-10.897 y=-533.369 z=288.851 mm, rx=-1.2337 ry=1.1953 rz=-1.2073 rad; joints [-51.497, -119.089, -83.078, -158.276, 37.645, 1.224] deg
          MoveL speed 250 mm/s, acceleration 1200 mm/s^2 (useActiveTCP=true optimoveEnabled=false optiMoveSpeed=0.3 optiMoveAcceleration=0.09) feature=Base
            Waypoint PosC_up: motionParameters(blendRadius=0.01); TCP in base x=241.567 y=-359.249 z=230.261 mm, rx=-1.2337 ry=1.1953 rz=-1.2073 rad; joints [-22.674, -126.16, -80.875, -153.323, 66.473, 0.967] deg
            Waypoint PosC_pick: motionParameters(jointSpeed=1.047198 jointAcceleration=1.396263 cartesianSpeed=0.05 cartesianAcceleration=0.3); TCP in base x=240.634 y=-361.553 z=93.98 mm, rx=-1.2337 ry=1.1953 rz=-1.2073 rad; joints [-22.914, -136.71, -85.338, -138.313, 66.273, 0.981] deg
            URCap Gripper (Robotiq_Grippers, Robotiq Inc.) dataModel(position=0.0, force=30.19607843137255, speed=30.19607843137255, positionInDouble=0.0, forceInDouble=30.19607843137255, speedInDouble=30.19607843137255, slaveIds=[9], blocking=true, robotCompliant=false)
            Waypoint PosC_up: TCP in base x=241.567 y=-359.249 z=230.261 mm, rx=-1.2337 ry=1.1953 rz=-1.2073 rad; joints [-22.674, -126.16, -80.875, -153.323, 66.473, 0.967] deg
            Waypoint Postions_otw: TCP in base x=-10.897 y=-533.369 z=288.851 mm, rx=-1.2337 ry=1.1953 rz=-1.2073 rad; joints [-51.497, -119.089, -83.078, -158.276, 37.645, 1.224] deg
          SafeHome (positionOptionType=SPEED_AND_ACCELERATION speed=1.047198 acceleration=1.396263 nextMotionTime=2)
          Num_cont_picked := Num_cont_picked+1
    Case (caseValue=48)
      Folder QR detections
        Device_ID := 1
        MoveJ speed 60 deg/s, acceleration 80 deg/s^2 (useActiveTCP=true optimoveEnabled=false optiMoveSpeed=0.3 optiMoveAcceleration=0.09) feature=Base
          Waypoint Variable (Variable): variable(featureName=Position1)
        URCap VISOR Trigger (SensoPart VISOR Robotic, SensoPart Industriesensorik GmbH) dataModel(visorId=0, visorSetJob=true, visorJobName=QR detection, visorImageAcqSetup=1); state(isChildrenLocked=true)
        pos1_powder := visor_getResponse(Device_ID)
        Script: pos1_powder = extract_powder_name(pos1_powder)
        MoveJ speed 60 deg/s, acceleration 80 deg/s^2 (useActiveTCP=true optimoveEnabled=false optiMoveSpeed=0.3 optiMoveAcceleration=0.09) feature=Base
          Waypoint Variable (Variable): variable(featureName=Position2)
        URCap VISOR Trigger (SensoPart VISOR Robotic, SensoPart Industriesensorik GmbH) dataModel(visorId=0, visorSetJob=true, visorJobName=QR detection, visorImageAcqSetup=1); state(isChildrenLocked=true)
        pos2_powder := visor_getResponse(Device_ID)
        Script: pos2_powder = extract_powder_name(pos2_powder)
        MoveJ speed 60 deg/s, acceleration 80 deg/s^2 (useActiveTCP=true optimoveEnabled=false optiMoveSpeed=0.3 optiMoveAcceleration=0.09) feature=Base
          Waypoint Variable (Variable): variable(featureName=Position3)
        URCap VISOR Trigger (SensoPart VISOR Robotic, SensoPart Industriesensorik GmbH) dataModel(visorId=0, visorSetJob=true, visorJobName=QR detection, visorImageAcqSetup=1); state(isChildrenLocked=true)
        pos3_powder := visor_getResponse(Device_ID)
        Script: pos3_powder = extract_powder_name(pos3_powder)
  '=========='
  Folder PostSettings [hidden by the author, left out]
